FUNCTION_BLOCK fbShutterAct
VAR

	OpenRelay : iRelay;
	CloseRelay : iRelay;
	
	CmdOpen : BOOL;
	CmdClose : BOOL;
	
	Config : stShutterConfig;
	StateType : eShutterStateType;
	
	OutputCheckTimer : TON;
END_VAR
VAR_OUTPUT
	Position : stShutterPosition;
END_VAR
VAR CONSTANT
	OutputCheckCycleTime: TIME := T#50MS;
END_VAR
VAR PERSISTENT
	HeightTime: TIME := T#0S;
	AngleTime: TIME := T#0S;
END_VAR


// Both signals must not be set at the same time
IF CmdOpen AND CmdClose THEN
	CmdOpen := FALSE;
	CmdClose := FALSE;
END_IF

// Reset signal if shutter reached fully open position with overstep
IF CmdOpen AND HeightTime >= Config.HeightTravelTime + Config.HeightTravelTimeOverstep THEN
	CmdOpen := FALSE;
END_IF

// Reset signal if shutter reached fully close position
IF CmdClose AND HeightTime <= T#0S THEN
	CmdClose := FALSE;
END_IF

// Write physical outputs and update shutter state
IF CmdOpen AND NOT CmdClose THEN
    CloseRelay.Reset();
    OpenRelay.Set();
	StateType := eShutterStateType.MOVING_UP;
ELSIF CmdClose AND NOT CmdOpen THEN
    OpenRelay.Reset();
    CloseRelay.Set();
	StateType := eShutterStateType.MOVING_DOWN;
ELSE
    OpenRelay.Reset();
    CloseRelay.Reset();
	StateType := eShutterStateType.IDLE;
END_IF

// Count time and accumulate when signals are set
OutputCheckTimer(IN := CmdOpen OR CmdClose, PT := OutputCheckCycleTime);
IF OutputCheckTimer.Q THEN
	IF CmdOpen THEN
		// Open fins first before moving up
		IF AngleTime < Config.AngleTravelTime THEN
			AngleTime := AngleTime + OutputCheckCycleTime;
		ELSIF HeightTime < Config.HeightTravelTime THEN
			HeightTime := HeightTime + OutputCheckCycleTime;
		END_IF;
	END_IF
	
	IF CmdClose THEN
		// Close fins first before moving down
		IF AngleTime > T#0S THEN
			AngleTime := AngleTime - OutputCheckCycleTime;
		ELSIF HeightTime > T#0s THEN
			HeightTime := HeightTime - OutputCheckCycleTime;
		END_IF;
	END_IF
	
	OutputCheckTimer.IN := FALSE;  // reset
END_IF

// Update shutter position% basen on position time
Position.Height := TimeToPosition(CurrentPosTime := HeightTime, TravelTime := Config.HeightTravelTime);
Position.Angle := TimeToPosition(CurrentPosTime := AngleTime, TravelTime := Config.AngleTravelTime);

METHOD Close
CmdOpen := FALSE;
CmdClose := TRUE;
END_METHOD

PROPERTY PUBLIC CurrentStateType : eShutterStateType
GET
CurrentStateType := This^.StateType;
END_GET
END_PROPERTY

//FB_Init is always available implicitly and it is used primarily for initialization.
//The return value is not evaluated. For a specific influence, you can also declare the
//methods explicitly and provide additional code there with the standard initialization
//code. You can evaluate the return value.
METHOD FB_Init: BOOL
VAR_INPUT
    bInitRetains: BOOL; // TRUE: the retain variables are initialized (reset warm / reset cold)
    bInCopyCode: BOOL;  // TRUE: the instance will be copied to the copy code afterward (online change)   
	
	OpenRelay : iRelay;
	CloseRelay : iRelay;
	Config : stShutterConfig;
	
END_VAR
THIS^.Config := Config;
THIS^.OpenRelay := OpenRelay;
THIS^.CloseRelay := CloseRelay;
END_METHOD

METHOD Open
CmdClose := FALSE;
CmdOpen := TRUE;
END_METHOD

METHOD Stop
CmdOpen := FALSE;
CmdClose := FALSE;
END_METHOD

METHOD PUBLIC TimeToPosition : USINT
VAR_INPUT
	CurrentPosTime : TIME;
	TravelTime : TIME;
END_VAR
IF TravelTime <= T#0S THEN
    TimeToPosition := 0;
ELSE
    TimeToPosition := UDINT_TO_USINT(100 * TIME_TO_UDINT(CurrentPosTime) / TIME_TO_UDINT(TravelTime));
END_IF
END_METHOD

END_FUNCTION_BLOCK

(* stored: Version 1.1.0.1
   POU fbShutterAct: Id {1ba23f45-b0eb-421e-9a3b-6a879c5afe8f}, SpecialFunc None
   Method Close: Id {f613d1a9-dcd5-4ce8-bd35-546352718445}
   Property CurrentStateType: Id {f29a13f8-1fef-4c57-98e7-dae28f0d5337}
   Get Get: Id {4ce8aa33-4386-4ae1-b83b-8847cdd706ea}
   Method FB_Init: Id {b49b88c3-5666-46b7-801a-0e8419ae9ce0}
   Method Open: Id {1dda91e8-cd15-4a31-9096-5e1a4c5f89a9}
   Method Stop: Id {17cc93a3-e742-4197-a775-db53f236a55d}
   Method TimeToPosition: Id {772cedc8-24ef-4e71-897a-f0415c3ffac2} *)
